(* Logix 5000 project; controller MECO9497 vendor 1 type 14 code 106 rev 21.11; software revision 21.00; part 3 of 4 *)
(* tags used below, declared in another part *)
   AAH_200 : BOOL;
   AAH_200_AUX : BOOL;
   AAH_200_DELAY : TIMER;
   ALARM_HORN_DO : ALIAS FOR Local:2:O.Data.10;
   ALARM_SCREEN_DISPLAY_BIT : BOOL;
   ALARM_SCREEN_LATCH_BIT : BOOL;
   ALERT_ALARM_SU_DELAY : TIMER;
   AT_200_AI : ALIAS FOR Local:4:I.Ch0Data;
   AT_200_EU : REAL;
   AUDIBLE_SUMMARY : BOOL;
   COMP_AMP_ALRM_DELAY_TMR : TIMER;
   COMPRESSOR_FAULT_DELAY : TIMER;
   COMPRESSOR_MOTOR_FLT_STARTUP_DELAY : TIMER;
   COMPRESSOR_MOTOR_START_DELAY : TIMER;
   COMPRESSOR_MOTOR_START_DO : ALIAS FOR Local:2:O.Data.0;
   COMPRESSOR_START_CMD : BOOL;
   CR_4 : ALIAS FOR Local:2:O.Data.9;
   CR_6 : ALIAS FOR Local:2:O.Data.2;
   CURRENT_SCREEN : DINT;
   D_V_REMOTE_START_MAP : BOOL;
   DIST_COND_ALRM_STARTUP_TMR : TIMER;
   DIST_PUMP_START_SP : REAL;
   DIST_PUMP_STOP_SP : REAL;
   DISTILLATE_MOTOR_FAULT_DELAY : TIMER;
   DISTILLATE_MOTOR_START_DO : ALIAS FOR Local:2:O.Data.1;
   DISTILLATE_PUMP_NORM_START : BOOL;
   DISTILLATE_PUMP_START_CMD : BOOL;
   DSTLT_BOX_DRAIN_NORM_DELAY : TIMER;
   DSTLT_PUMP_START_DELAY : TIMER;
   DSTLT_STORAGE : BOOL;
   DSTLT_STORAGE_DELAY_TIMER : TIMER;
   DSTLT_STORAGE_ENABLE_MAP : BOOL;
   DSTLT_TEMP_ALRM_SU_DELAY : TIMER;
   DSTLT_TEMP_CNTRL_DELAY_TIMER : TIMER;
   E_Stop_AUX : BOOL;
   ENGINEER : BOOL;
   EVAP_PRESSURE_PERM : BOOL;
   EVAP_PRESSURE_PERM_TIMER : TIMER;
   EVAP_RAMP_ENABLE_DELAY_TIMER : TIMER;
   EXCESS_DIST_TO_DRAIN_AUX : BOOL;
   EXCESS_DSTLT_DELAY_TIMER : TIMER;
   EXCESS_DSTLT_DRAIN : BOOL;
   EXCESS_DSTLT_DRAIN_TIMER : TIMER;
   EXCESS_DSTLT_REMAIN : DINT;
   FC_300_AM_OIT : BOOL;
   FC_300_SP : DINT;
   FC_300_SP_OUT : DINT;
   FT_200_AI : ALIAS FOR Local:3:I.Ch2Data;
   FT_200_EU : REAL;
   HEARTBEAT_AUX : BOOL;
   HOT_STANDBY : BOOL;
   HOURMETER_DO : ALIAS FOR Local:2:O.Data.4;
   IAL_100_AUX : BOOL;
   INITIAL_SCAN_BIT : BOOL;
   INITIAL_SCAN_SYS_RESET : BOOL;
   INITIAL_SCAN_SYS_RESET_TMR : TIMER;
   IY_100_AI : ALIAS FOR Local:4:I.Ch2Data;
   IY_100_EU : REAL;
   LAH_100_AUX : BOOL;
   LAL_100_AUX : BOOL;
   LB_OIL_LOW_PRESS_ALRM_DELAY : TIMER;
   LCV_100_IND : DINT;
   LCV_200_IND : DINT;
   LIC_100 : PID;
   LIC_200 : PID;
   LT_100_AI : ALIAS FOR Local:3:I.Ch3Data;
   LT_100_EU : REAL;
   LT_200_AI : ALIAS FOR Local:3:I.Ch4Data;
   LT_200_EU : REAL;
   LUBE_OIL_PUMP_FAULT_DELAY : TIMER;
   LUBE_OIL_PUMP_START_CMD : BOOL;
   LUBE_OIL_SHUTDWN_TIMER : TIMER;
   M1_DI_MAP : BOOL;
   M1_FAULT_AUX : BOOL;
   M2_DI_MAP : BOOL;
   M2_FAULT_AUX : BOOL;
   M4_DI_MAP : BOOL;
   M4_FAULT_AUX : BOOL;
   MAINTENANCE : BOOL;
   MCB : BOOL;
   MSG_AAH_200 : BOOL;
   MSG_E_STOP : BOOL;
   MSG_EXCESS_DIST_TO_DRAIN : BOOL;
   MSG_IAL_100 : BOOL;
   MSG_LAH_100 : BOOL;
   MSG_LAL_100 : BOOL;
   MSG_M1_FLT : BOOL;
   MSG_M2_FLT : BOOL;
   MSG_M4_FLT : BOOL;
   MSG_PAH_103 : BOOL;
   MSG_PAL_103 : BOOL;
   MSG_PAL_700 : BOOL;
   MSG_TAH_700 : BOOL;
   MSG_TAL_200 : BOOL;
   MSS_SHUTDOWN : BOOL;
   MSS_START_PERM : BOOL;
   OIL_MOTOR_START_DO : ALIAS FOR Local:2:O.Data.11;
   OIT_SCREEN_CONTROL : DINT;
   OIT_SECURITY_LEVEL : DINT;
   OP_SWTCH_AUTO_DI_MAP : BOOL;
   OP_SWTCH_MANUAL_DI_MAP : BOOL;
   OPERATOR : BOOL;
   PAH_103_AUX : BOOL;
   PAL_103_AUX : BOOL;
   PAL_700_AUX : BOOL;
   PCV_103_IND : DINT;
   PERM_TIME_REMAINING : REAL;
   PIC_103 : PID;
   PT_103_AI : ALIAS FOR Local:3:I.Ch0Data;
   PT_103_EU : REAL;
   SECURITY_ENABLED : BOOL;
   SV_200 : ALIAS FOR Local:2:O.Data.5;
   SV_200_201_DO : ALIAS FOR Local:2:O.Data.6;
   SV_200_201_IND : BOOL;
   SV_200_CTL : BOOL;
   SV_200_IND : BOOL;
   SV_500_DO : ALIAS FOR Local:2:O.Data.8;
   SV_500_IND : BOOL;
   TAH_700_AUX : BOOL;
   TAL_200 : BOOL;
   TAL_200_AUX : BOOL;
   TAL_200_DELAY : TIMER;
   TCV_102_IND : DINT;
   TCV_200_IND : DINT;
   TIC_102 : PID;
   TIC_200 : PID;
   TT_102_AI : ALIAS FOR Local:3:I.Ch1Data;
   TT_102_EU : REAL;
   TT_200_AI : ALIAS FOR Local:4:I.Ch1Data;
   TT_200_EU : REAL;
   UNIT_REMOTE_START_MAP : BOOL;
   UNIT_START_DI_MAP : BOOL;
   UNIT_STATUS : DINT;
   UNIT_STOP_DI_MAP : BOOL;
(* MainProgram, continued *)

ROUTINE MainRoutine   (* ladder *)
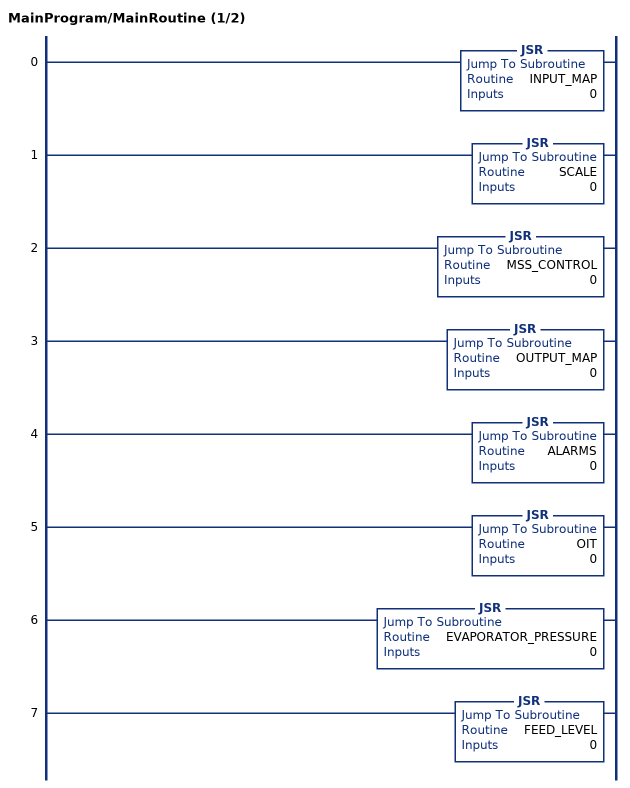
   0: JSR(INPUT_MAP,0);
   1: JSR(SCALE,0);
   2: JSR(MSS_CONTROL,0);
   3: JSR(OUTPUT_MAP,0);
   4: JSR(ALARMS,0);
   5: JSR(OIT,0);
   6: JSR(EVAPORATOR_PRESSURE,0);
   7: JSR(FEED_LEVEL,0);
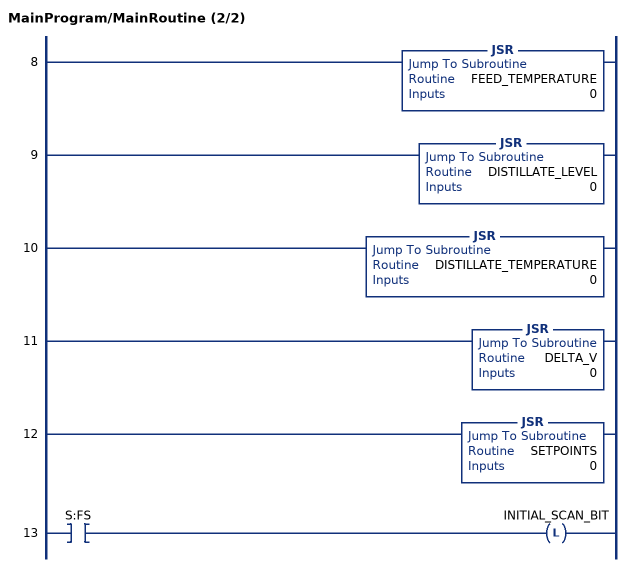
   8: JSR(FEED_TEMPERATURE,0);
   9: JSR(DISTILLATE_LEVEL,0);
   10: JSR(DISTILLATE_TEMPERATURE,0);
   11: JSR(DELTA_V,0);
   12: JSR(SETPOINTS,0);
   13: XIC(S:FS)OTL(INITIAL_SCAN_BIT);
END_ROUTINE

ROUTINE MSS_CONTROL   (* ladder *)
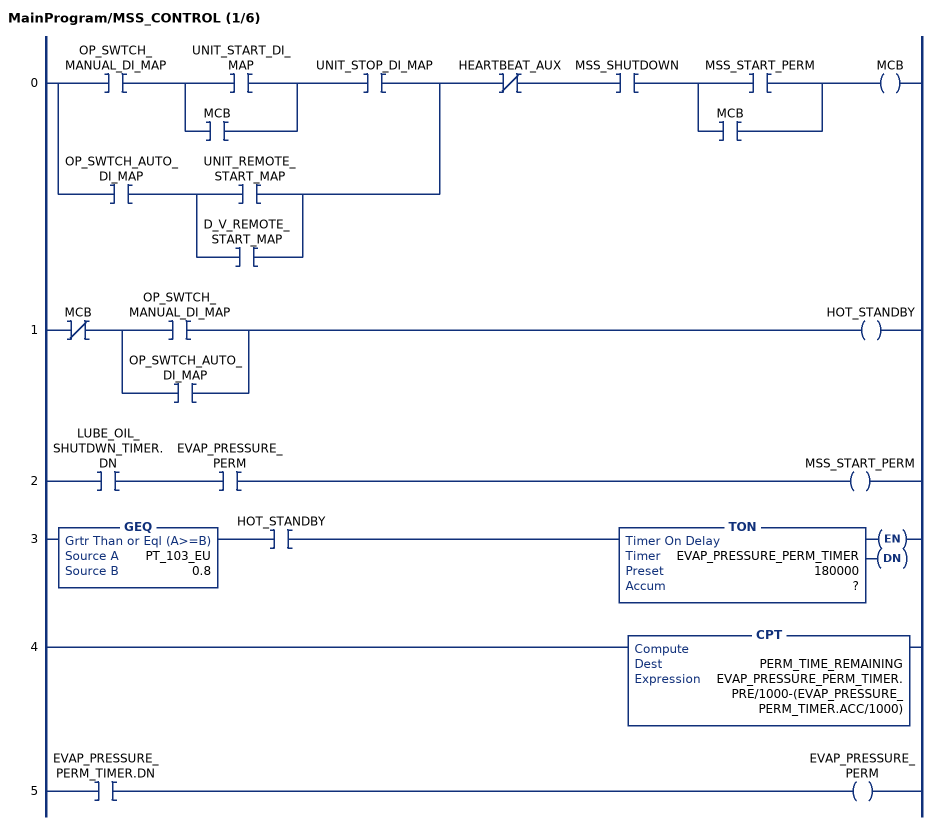
   0: [XIC(OP_SWTCH_MANUAL_DI_MAP) [XIC(UNIT_START_DI_MAP) ,XIC(MCB) ] XIC(UNIT_STOP_DI_MAP) ,XIC(OP_SWTCH_AUTO_DI_MAP) [XIC(UNIT_REMOTE_START_MAP) ,XIC(D_V_REMOTE_START_MAP) ] ]XIO(HEARTBEAT_AUX)XIC(MSS_SHUTDOWN)[XIC(MSS_START_PERM) ,XIC(MCB) ]OTE(MCB);
   1: XIO(MCB)[XIC(OP_SWTCH_MANUAL_DI_MAP) ,XIC(OP_SWTCH_AUTO_DI_MAP) ]OTE(HOT_STANDBY);
   2: XIC(LUBE_OIL_SHUTDWN_TIMER.DN)XIC(EVAP_PRESSURE_PERM)OTE(MSS_START_PERM);
   3: GEQ(PT_103_EU,0.8)XIC(HOT_STANDBY)TON(EVAP_PRESSURE_PERM_TIMER,?,?);
   4: CPT(PERM_TIME_REMAINING,EVAP_PRESSURE_PERM_TIMER.PRE/1000-(EVAP_PRESSURE_PERM_TIMER.ACC/1000));
   5: XIC(EVAP_PRESSURE_PERM_TIMER.DN)OTE(EVAP_PRESSURE_PERM);
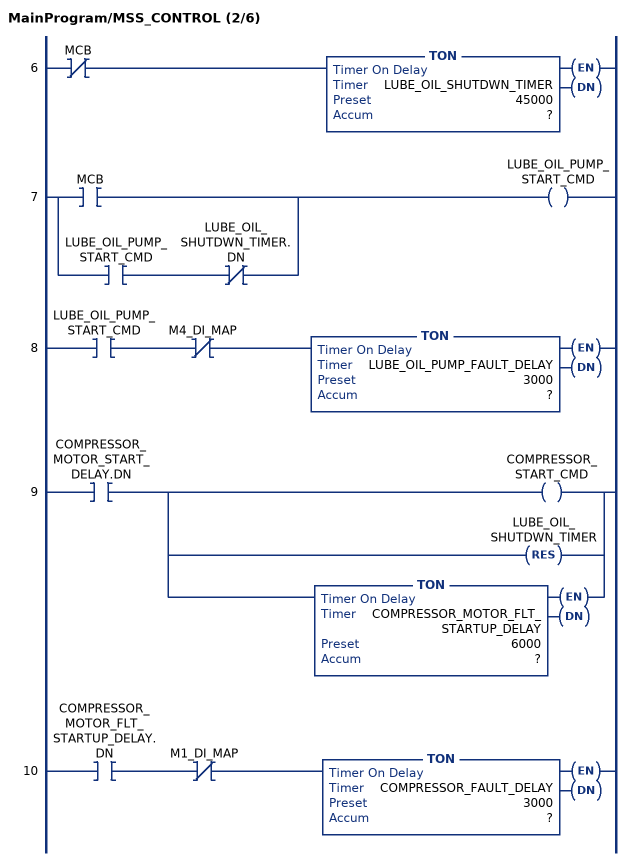
   6: XIO(MCB)TON(LUBE_OIL_SHUTDWN_TIMER,?,?);
   7: [XIC(MCB) ,XIC(LUBE_OIL_PUMP_START_CMD) XIO(LUBE_OIL_SHUTDWN_TIMER.DN) ]OTE(LUBE_OIL_PUMP_START_CMD);
   8: XIC(LUBE_OIL_PUMP_START_CMD)XIO(M4_DI_MAP)TON(LUBE_OIL_PUMP_FAULT_DELAY,?,?);
   9: XIC(COMPRESSOR_MOTOR_START_DELAY.DN)[OTE(COMPRESSOR_START_CMD) ,RES(LUBE_OIL_SHUTDWN_TIMER) ,TON(COMPRESSOR_MOTOR_FLT_STARTUP_DELAY,?,?) ];
   10: XIC(COMPRESSOR_MOTOR_FLT_STARTUP_DELAY.DN)XIO(M1_DI_MAP)TON(COMPRESSOR_FAULT_DELAY,?,?);
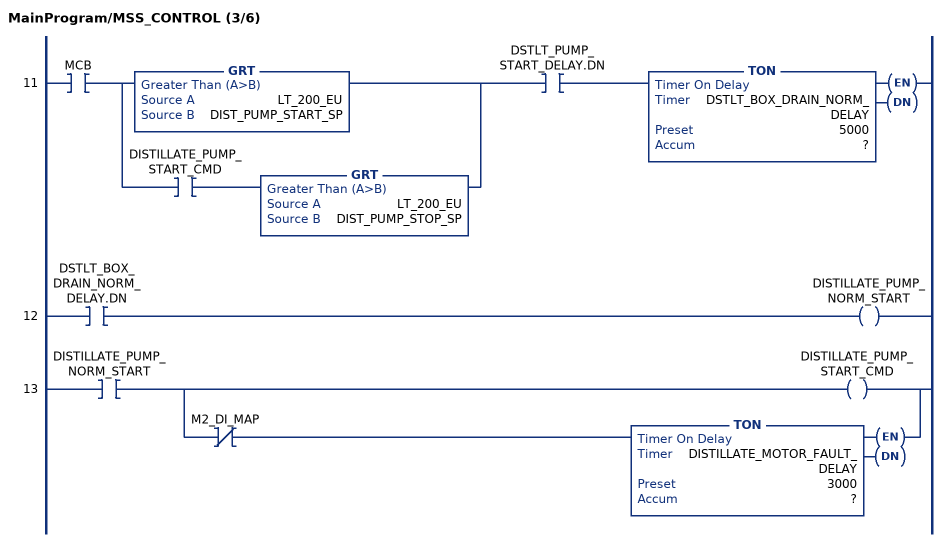
   11: XIC(MCB)[GRT(LT_200_EU,DIST_PUMP_START_SP) ,XIC(DISTILLATE_PUMP_START_CMD) GRT(LT_200_EU,DIST_PUMP_STOP_SP) ]XIC(DSTLT_PUMP_START_DELAY.DN)TON(DSTLT_BOX_DRAIN_NORM_DELAY,?,?);
   12: XIC(DSTLT_BOX_DRAIN_NORM_DELAY.DN)OTE(DISTILLATE_PUMP_NORM_START);
   13: XIC(DISTILLATE_PUMP_NORM_START)[OTE(DISTILLATE_PUMP_START_CMD) ,XIO(M2_DI_MAP) TON(DISTILLATE_MOTOR_FAULT_DELAY,?,?) ];
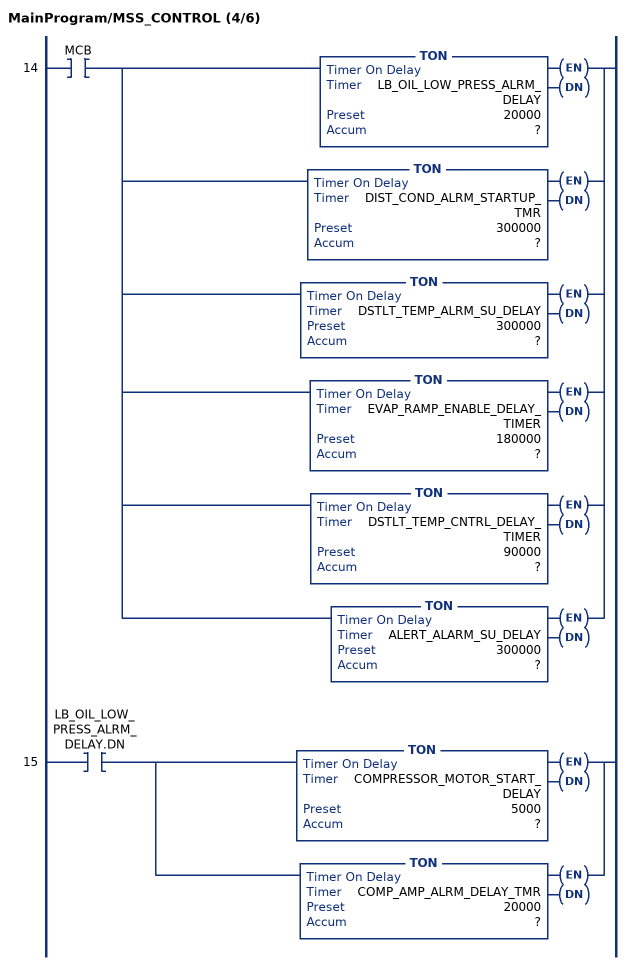
   14: XIC(MCB)[TON(LB_OIL_LOW_PRESS_ALRM_DELAY,?,?) ,TON(DIST_COND_ALRM_STARTUP_TMR,?,?) ,TON(DSTLT_TEMP_ALRM_SU_DELAY,?,?) ,TON(EVAP_RAMP_ENABLE_DELAY_TIMER,?,?) ,TON(DSTLT_TEMP_CNTRL_DELAY_TIMER,?,?) ,TON(ALERT_ALARM_SU_DELAY,?,?) ];
   15: XIC(LB_OIL_LOW_PRESS_ALRM_DELAY.DN)[TON(COMPRESSOR_MOTOR_START_DELAY,?,?) ,TON(COMP_AMP_ALRM_DELAY_TMR,?,?) ];
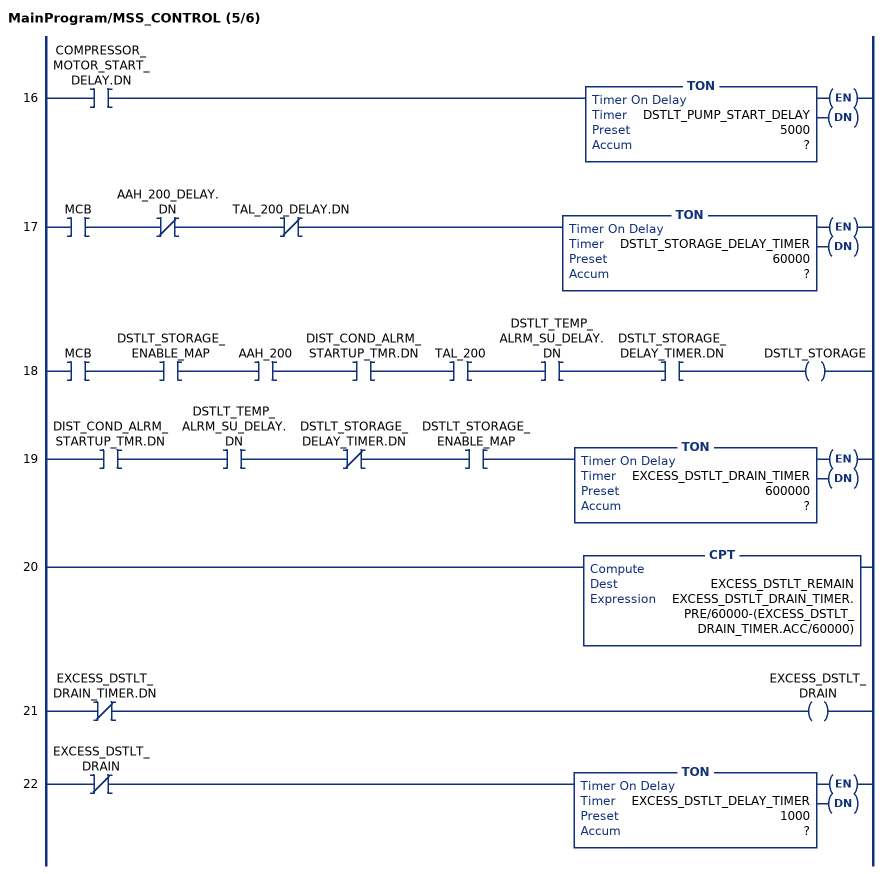
   16: XIC(COMPRESSOR_MOTOR_START_DELAY.DN)TON(DSTLT_PUMP_START_DELAY,?,?);
   17: XIC(MCB)XIO(AAH_200_DELAY.DN)XIO(TAL_200_DELAY.DN)TON(DSTLT_STORAGE_DELAY_TIMER,?,?);
   18: XIC(MCB)XIC(DSTLT_STORAGE_ENABLE_MAP)XIC(AAH_200)XIC(DIST_COND_ALRM_STARTUP_TMR.DN)XIC(TAL_200)XIC(DSTLT_TEMP_ALRM_SU_DELAY.DN)XIC(DSTLT_STORAGE_DELAY_TIMER.DN)OTE(DSTLT_STORAGE);
   19: XIC(DIST_COND_ALRM_STARTUP_TMR.DN)XIC(DSTLT_TEMP_ALRM_SU_DELAY.DN)XIO(DSTLT_STORAGE_DELAY_TIMER.DN)XIC(DSTLT_STORAGE_ENABLE_MAP)TON(EXCESS_DSTLT_DRAIN_TIMER,?,?);
   20: CPT(EXCESS_DSTLT_REMAIN,EXCESS_DSTLT_DRAIN_TIMER.PRE/60000-(EXCESS_DSTLT_DRAIN_TIMER.ACC/60000));
   21: XIO(EXCESS_DSTLT_DRAIN_TIMER.DN)OTE(EXCESS_DSTLT_DRAIN);
   22: XIO(EXCESS_DSTLT_DRAIN)TON(EXCESS_DSTLT_DELAY_TIMER,?,?);
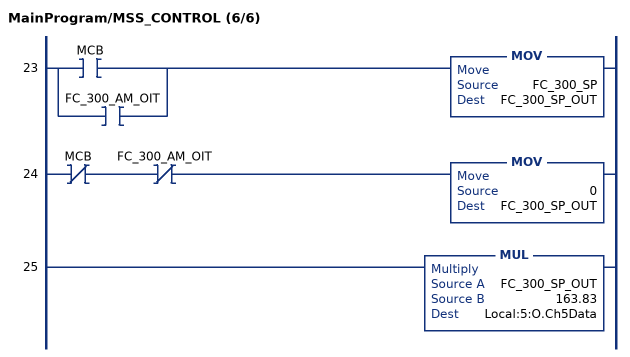
   23: [XIC(MCB) ,XIC(FC_300_AM_OIT) ]MOV(FC_300_SP,FC_300_SP_OUT);
   24: XIO(MCB)XIO(FC_300_AM_OIT)MOV(0,FC_300_SP_OUT);
   25: MUL(FC_300_SP_OUT,163.83,Local:5:O.Ch5Data);
END_ROUTINE

ROUTINE OIT   (* ladder *)
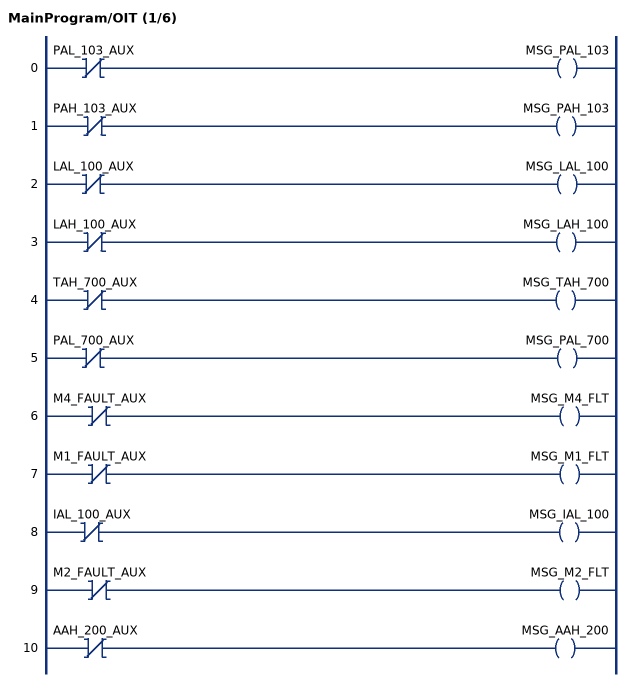
   0: XIO(PAL_103_AUX)OTE(MSG_PAL_103);
   1: XIO(PAH_103_AUX)OTE(MSG_PAH_103);
   2: XIO(LAL_100_AUX)OTE(MSG_LAL_100);
   3: XIO(LAH_100_AUX)OTE(MSG_LAH_100);
   4: XIO(TAH_700_AUX)OTE(MSG_TAH_700);
   5: XIO(PAL_700_AUX)OTE(MSG_PAL_700);
   6: XIO(M4_FAULT_AUX)OTE(MSG_M4_FLT);
   7: XIO(M1_FAULT_AUX)OTE(MSG_M1_FLT);
   8: XIO(IAL_100_AUX)OTE(MSG_IAL_100);
   9: XIO(M2_FAULT_AUX)OTE(MSG_M2_FLT);
   10: XIO(AAH_200_AUX)OTE(MSG_AAH_200);
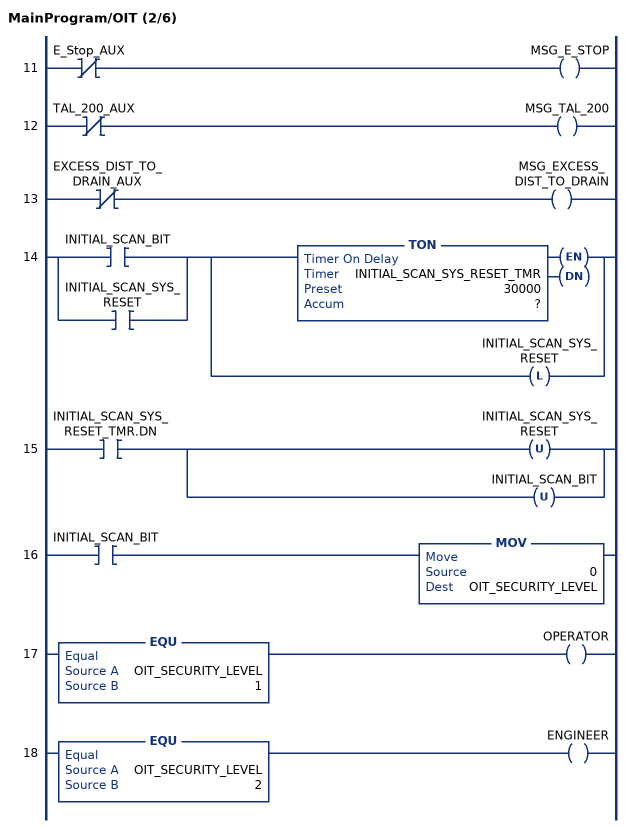
   11: XIO(E_Stop_AUX)OTE(MSG_E_STOP);
   12: XIO(TAL_200_AUX)OTE(MSG_TAL_200);
   13: XIO(EXCESS_DIST_TO_DRAIN_AUX)OTE(MSG_EXCESS_DIST_TO_DRAIN);
   14: [XIC(INITIAL_SCAN_BIT) ,XIC(INITIAL_SCAN_SYS_RESET) ][TON(INITIAL_SCAN_SYS_RESET_TMR,?,?) ,OTL(INITIAL_SCAN_SYS_RESET) ];
   15: XIC(INITIAL_SCAN_SYS_RESET_TMR.DN)[OTU(INITIAL_SCAN_SYS_RESET) ,OTU(INITIAL_SCAN_BIT) ];
   16: XIC(INITIAL_SCAN_BIT)MOV(0,OIT_SECURITY_LEVEL);
   17: EQU(OIT_SECURITY_LEVEL,1)OTE(OPERATOR);
   18: EQU(OIT_SECURITY_LEVEL,2)OTE(ENGINEER);
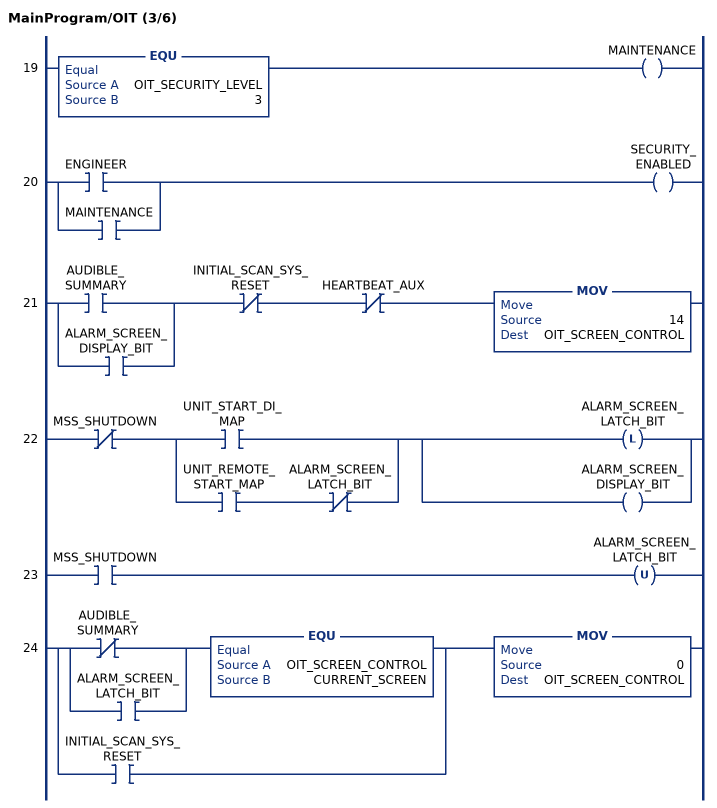
   19: EQU(OIT_SECURITY_LEVEL,3)OTE(MAINTENANCE);
   20: [XIC(ENGINEER) ,XIC(MAINTENANCE) ]OTE(SECURITY_ENABLED);
   21: [XIC(AUDIBLE_SUMMARY) ,XIC(ALARM_SCREEN_DISPLAY_BIT) ]XIO(INITIAL_SCAN_SYS_RESET)XIO(HEARTBEAT_AUX)MOV(14,OIT_SCREEN_CONTROL);
   22: XIO(MSS_SHUTDOWN)[XIC(UNIT_START_DI_MAP) ,XIC(UNIT_REMOTE_START_MAP) XIO(ALARM_SCREEN_LATCH_BIT) ][OTL(ALARM_SCREEN_LATCH_BIT) ,OTE(ALARM_SCREEN_DISPLAY_BIT) ];
   23: XIC(MSS_SHUTDOWN)OTU(ALARM_SCREEN_LATCH_BIT);
   24: [[XIO(AUDIBLE_SUMMARY) ,XIC(ALARM_SCREEN_LATCH_BIT) ] EQU(OIT_SCREEN_CONTROL,CURRENT_SCREEN) ,XIC(INITIAL_SCAN_SYS_RESET) ]MOV(0,OIT_SCREEN_CONTROL);
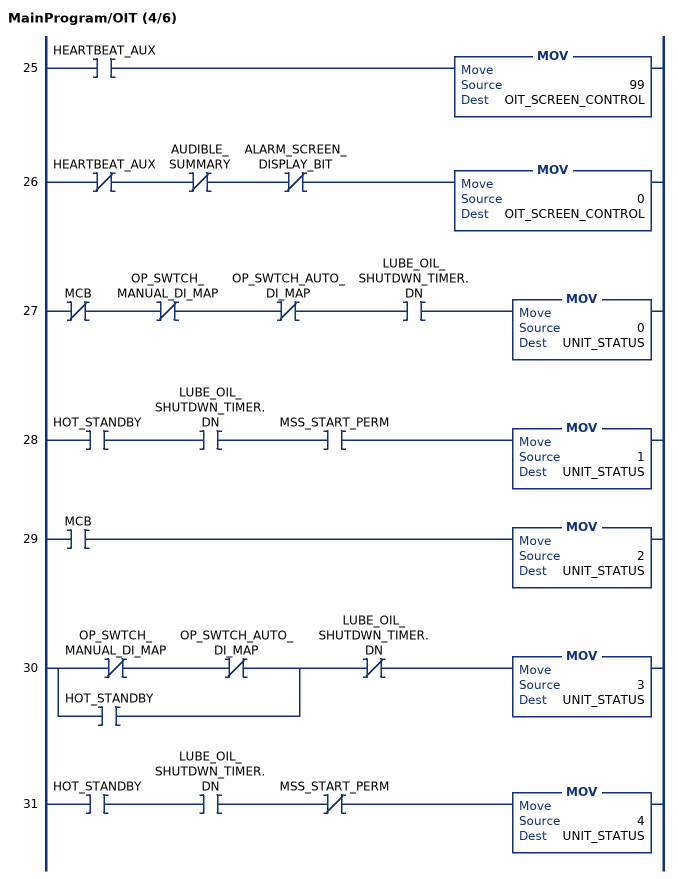
   25: XIC(HEARTBEAT_AUX)MOV(99,OIT_SCREEN_CONTROL);
   26: XIO(HEARTBEAT_AUX)XIO(AUDIBLE_SUMMARY)XIO(ALARM_SCREEN_DISPLAY_BIT)MOV(0,OIT_SCREEN_CONTROL);
   27: XIO(MCB)XIO(OP_SWTCH_MANUAL_DI_MAP)XIO(OP_SWTCH_AUTO_DI_MAP)XIC(LUBE_OIL_SHUTDWN_TIMER.DN)MOV(0,UNIT_STATUS);
   28: XIC(HOT_STANDBY)XIC(LUBE_OIL_SHUTDWN_TIMER.DN)XIC(MSS_START_PERM)MOV(1,UNIT_STATUS);
   29: XIC(MCB)MOV(2,UNIT_STATUS);
   30: [XIO(OP_SWTCH_MANUAL_DI_MAP) XIO(OP_SWTCH_AUTO_DI_MAP) ,XIC(HOT_STANDBY) ]XIO(LUBE_OIL_SHUTDWN_TIMER.DN)MOV(3,UNIT_STATUS);
   31: XIC(HOT_STANDBY)XIC(LUBE_OIL_SHUTDWN_TIMER.DN)XIO(MSS_START_PERM)MOV(4,UNIT_STATUS);
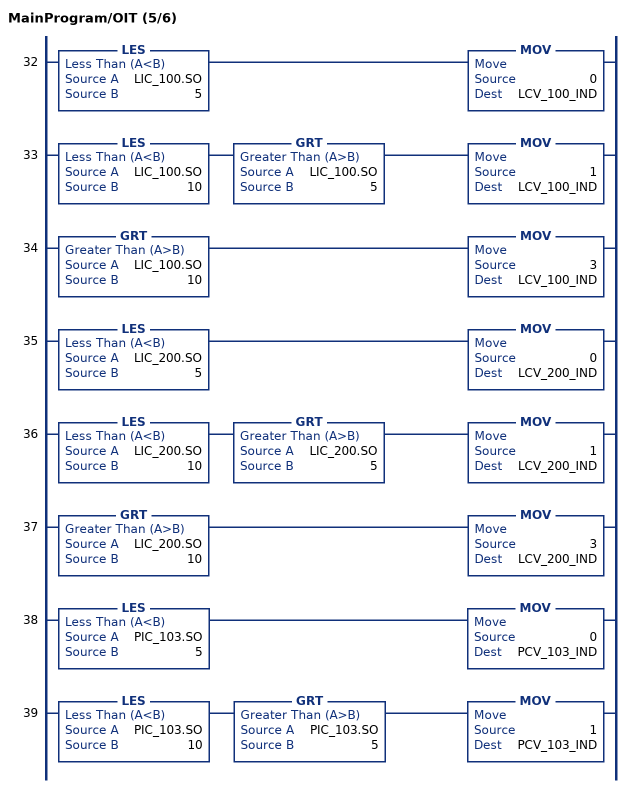
   32: LES(LIC_100.SO,5)MOV(0,LCV_100_IND);
   33: LES(LIC_100.SO,10)GRT(LIC_100.SO,5)MOV(1,LCV_100_IND);
   34: GRT(LIC_100.SO,10)MOV(3,LCV_100_IND);
   35: LES(LIC_200.SO,5)MOV(0,LCV_200_IND);
   36: LES(LIC_200.SO,10)GRT(LIC_200.SO,5)MOV(1,LCV_200_IND);
   37: GRT(LIC_200.SO,10)MOV(3,LCV_200_IND);
   38: LES(PIC_103.SO,5)MOV(0,PCV_103_IND);
   39: LES(PIC_103.SO,10)GRT(PIC_103.SO,5)MOV(1,PCV_103_IND);
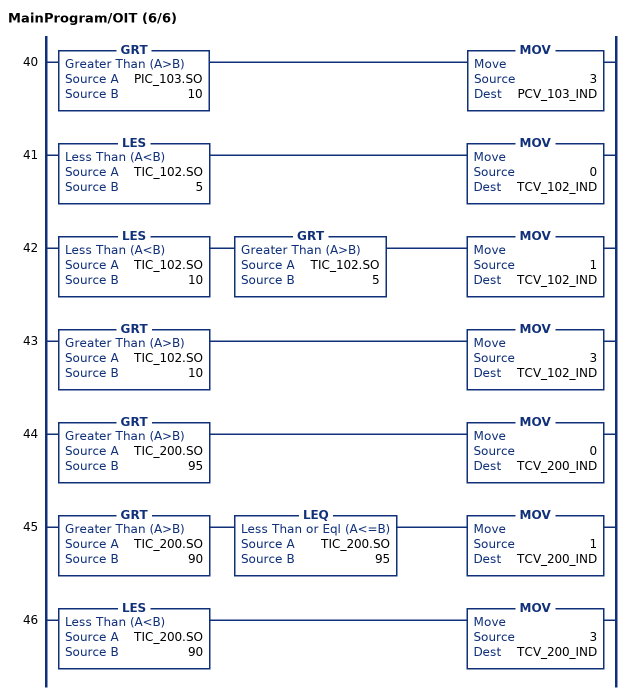
   40: GRT(PIC_103.SO,10)MOV(3,PCV_103_IND);
   41: LES(TIC_102.SO,5)MOV(0,TCV_102_IND);
   42: LES(TIC_102.SO,10)GRT(TIC_102.SO,5)MOV(1,TCV_102_IND);
   43: GRT(TIC_102.SO,10)MOV(3,TCV_102_IND);
   44: GRT(TIC_200.SO,95)MOV(0,TCV_200_IND);
   45: GRT(TIC_200.SO,90)LEQ(TIC_200.SO,95)MOV(1,TCV_200_IND);
   46: LES(TIC_200.SO,90)MOV(3,TCV_200_IND);
END_ROUTINE

ROUTINE OUTPUT_MAP   (* ladder *)
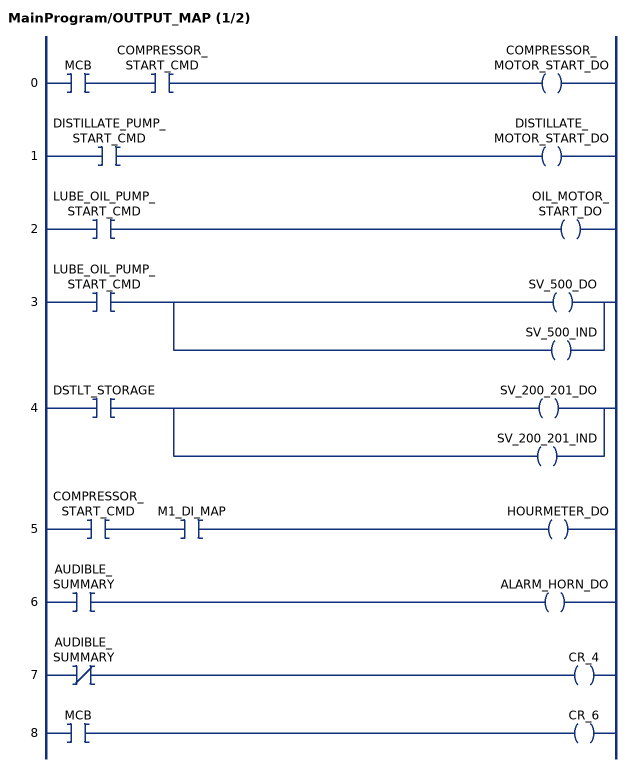
   0: XIC(MCB)XIC(COMPRESSOR_START_CMD)OTE(COMPRESSOR_MOTOR_START_DO);
   1: XIC(DISTILLATE_PUMP_START_CMD)OTE(DISTILLATE_MOTOR_START_DO);
   2: XIC(LUBE_OIL_PUMP_START_CMD)OTE(OIL_MOTOR_START_DO);
   3: XIC(LUBE_OIL_PUMP_START_CMD)[OTE(SV_500_DO) ,OTE(SV_500_IND) ];
   4: XIC(DSTLT_STORAGE)[OTE(SV_200_201_DO) ,OTE(SV_200_201_IND) ];
   5: XIC(COMPRESSOR_START_CMD)XIC(M1_DI_MAP)OTE(HOURMETER_DO);
   6: XIC(AUDIBLE_SUMMARY)OTE(ALARM_HORN_DO);
   7: XIO(AUDIBLE_SUMMARY)OTE(CR_4);
   8: XIC(MCB)OTE(CR_6);
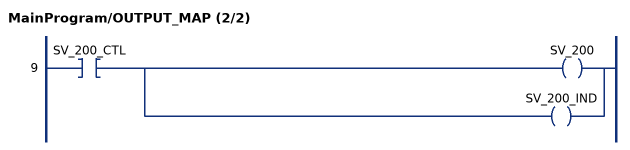
   9: XIC(SV_200_CTL)[OTE(SV_200) ,OTE(SV_200_IND) ];
END_ROUTINE

ROUTINE SCALE   (* function block diagram *)
   SHEET 1
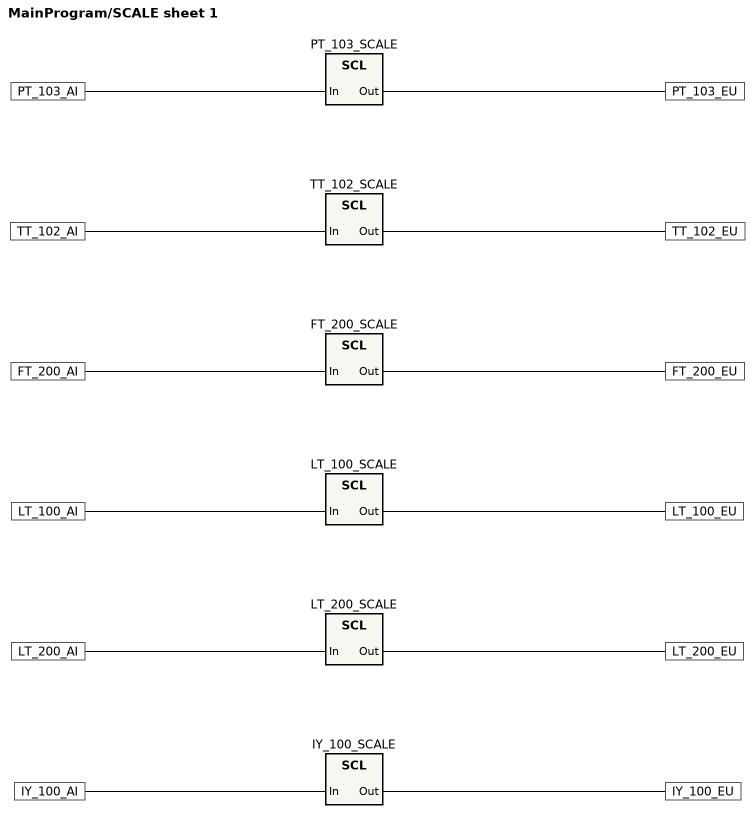
   PT_103_SCALE : SCL(In := PT_103_AI);
   TT_102_SCALE : SCL(In := TT_102_AI);
   FT_200_SCALE : SCL(In := FT_200_AI);
   LT_100_SCALE : SCL(In := LT_100_AI);
   LT_200_SCALE : SCL(In := LT_200_AI);
   IY_100_SCALE : SCL(In := IY_100_AI);
   PT_103_EU := PT_103_SCALE.Out;
   TT_102_EU := TT_102_SCALE.Out;
   FT_200_EU := FT_200_SCALE.Out;
   LT_100_EU := LT_100_SCALE.Out;
   LT_200_EU := LT_200_SCALE.Out;
   IY_100_EU := IY_100_SCALE.Out;
   SHEET 2
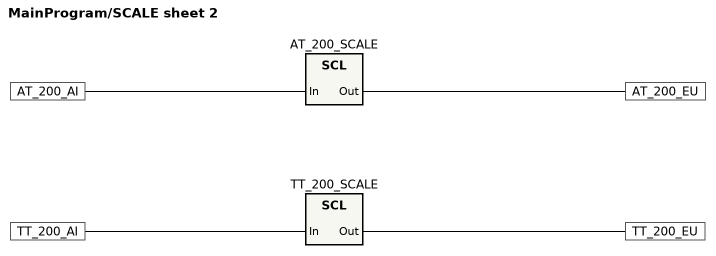
   AT_200_SCALE : SCL(In := AT_200_AI);
   TT_200_SCALE : SCL(In := TT_200_AI);
   AT_200_EU := AT_200_SCALE.Out;
   TT_200_EU := TT_200_SCALE.Out;
END_ROUTINE
